(* IEC 61131-3 sources: sps-foerderband-sortieranlage/plc, 10 files *)

(* ---- E_Schritt.st ---- *)
{attribute 'qualified_only'}
{attribute 'strict'}
TYPE E_Schritt :
(
    INIT            := 0,   // Grundstellung herstellen
    BEREIT          := 1,   // Stillstand, wartet auf Start
    WARTEN_AUF_TEIL := 2,   // Automatik, wartet auf Teil an B1
    TRANSPORT       := 3,   // Band läuft, Material wird an B2 erkannt
    AUSWERFER_AUS   := 4,   // Metallteil: Auswerfer fährt aus
    AUSWERFER_EIN   := 5,   // Auswerfer fährt zurück
    STOERUNG        := 9    // Not-Halt oder Zeitüberschreitung
);
END_TYPE

(* ---- GVL_IO.st ---- *)
{attribute 'qualified_only'}
VAR_GLOBAL
    // ---------- Eingänge ----------
    // Öffner: TRUE = in Ordnung. Startwert TRUE nur für die Simulation,
    // weil es keinen realen Taster gibt, der den Kontakt geschlossen hält.
    xNotHaltOk            : BOOL := TRUE;   // S0  %IX0.0  Öffner
    xStart                : BOOL;           // S1  %IX0.1  Schließer
    xStoppOk              : BOOL := TRUE;   // S2  %IX0.2  Öffner
    xQuittieren           : BOOL;           // S3  %IX0.3  Schließer
    xZaehlerReset         : BOOL;           // S4  %IX0.4  Schließer
    xTeilEinlauf          : BOOL;           // B1  %IX0.5
    xTeilMetall           : BOOL;           // B2  %IX0.6  induktiv
    xTeilAuswurfPos       : BOOL;           // B3  %IX0.7
    xTeilRutscheB         : BOOL;           // B4  %IX1.0
    xAuswerferEingefahren : BOOL := TRUE;   // B5  %IX1.1
    xAuswerferAusgefahren : BOOL;           // B6  %IX1.2

    // ---------- Ausgänge ----------
    xBandMotor            : BOOL;           // K1/M1 %QX0.0
    xAuswerferAusfahren   : BOOL;           // Y1    %QX0.1
    xLampeBetrieb         : BOOL;           // H1    %QX0.2
    xLampeStoerung        : BOOL;           // H2    %QX0.3
END_VAR

(* ---- GVL_Param.st ---- *)
{attribute 'qualified_only'}
VAR_GLOBAL CONSTANT
    tTimeoutTransport : TIME := T#8S;     // Teil muss B3 bzw. B4 innerhalb dieser Zeit erreichen
    tTimeoutAuswerfer : TIME := T#2S;     // Auswerfer muss seine Endlage innerhalb dieser Zeit erreichen
    tBlinkHalbperiode : TIME := T#500MS;  // Blinktakt der Störungsleuchte
END_VAR

(* ---- GVL_Sim.st ---- *)
{attribute 'qualified_only'}
VAR_GLOBAL
    // ---------- Bedienung der Simulation (Visualisierung) ----------
    xMetallteilAuflegen     : BOOL;
    xKunststoffteilAuflegen : BOOL;
    xBandLeeren             : BOOL;      // Bediener nimmt ein Teil vom Band (z. B. nach Not-Halt)
    xZylinderKlemmt         : BOOL;      // Fehlersimulation: Auswerfer bewegt sich nicht

    // ---------- Zustand der Simulation (nur Anzeige) ----------
    xTeilAufBand            : BOOL;
    rTeilPosition           : REAL;      // mm ab Bandanfang
    rAuswerferPosition      : REAL;      // 0 = eingefahren, 100 = ausgefahren
END_VAR

(* ---- GVL_Status.st ---- *)
{attribute 'qualified_only'}
VAR_GLOBAL
    // ---------- Zustand (wird per OPC UA bereitgestellt) ----------
    eSchritt            : E_Schritt := E_Schritt.INIT;
    sSchritt            : STRING(30);
    xBetrieb            : BOOL;          // Automatikablauf aktiv
    xStoerung           : BOOL;          // Störung gespeichert, noch nicht quittiert
    xNotHaltAktiv       : BOOL;          // Not-Halt steht aktuell an
    sStoerung           : STRING(80);    // Störungstext

    // ---------- Zähler und Kennzahlen ----------
    uiAnzahlMetall      : UINT;
    uiAnzahlKunststoff  : UINT;
    uiAnzahlGesamt      : UINT;
    uiAnzahlNotHalt     : UINT;
    tLetzteZykluszeit   : TIME;          // Zeit vom Einlauf bis zum Abschluss des letzten Teils
    tStillstandGesamt   : TIME;          // aufsummierte Zeit im Störungszustand

    // ---------- interne Anforderungen Ablauf -> Ausgaben ----------
    xBandEin            : BOOL;
    xAuswerferEin       : BOOL;
END_VAR

(* ---- FB_Anlagensimulation.st ---- *)
FUNCTION_BLOCK FB_Anlagensimulation
VAR
    fbMetallFlanke     : R_TRIG;
    fbKunststoffFlanke : R_TRIG;
    fbLeerenFlanke     : R_TRIG;
    fbRutscheBImpuls   : TP;
    xTeilIstMetall     : BOOL;
    xTeilFaelltInB     : BOOL;
    xErsterZyklus      : BOOL := TRUE;
    tJetzt             : TIME;
    tLetzter           : TIME;
    rDt                : REAL;          // Zeit seit dem letzten Zyklus in s
END_VAR
VAR CONSTANT
    rBandGeschw        : REAL := 200.0;  // mm/s
    rBandLaenge        : REAL := 1000.0; // mm
    rB1Start           : REAL := 0.0;
    rB1Ende            : REAL := 80.0;
    rB2Start           : REAL := 350.0;
    rB2Ende            : REAL := 420.0;
    rB3Start           : REAL := 650.0;
    rB3Ende            : REAL := 720.0;
    rAuswerferGeschw   : REAL := 200.0;  // %/s, ein Hub dauert 0,5 s
    rAuswurfSchwelle   : REAL := 50.0;   // ab hier ist das Teil vom Band geschoben
END_VAR

(* ---------- Implementierung ---------- *)

// Zeitschritt bestimmen (begrenzt, damit Pausen im Debugger keine Sprünge erzeugen)
tJetzt := TIME();
IF xErsterZyklus THEN
    tLetzter := tJetzt;
    xErsterZyklus := FALSE;
END_IF
rDt := MIN(TIME_TO_REAL(tJetzt - tLetzter) / 1000.0, 0.1);
tLetzter := tJetzt;

// Teile auflegen und entfernen
fbMetallFlanke(CLK := GVL_Sim.xMetallteilAuflegen);
fbKunststoffFlanke(CLK := GVL_Sim.xKunststoffteilAuflegen);
fbLeerenFlanke(CLK := GVL_Sim.xBandLeeren);

IF NOT GVL_Sim.xTeilAufBand THEN
    IF fbMetallFlanke.Q THEN
        GVL_Sim.xTeilAufBand := TRUE;
        GVL_Sim.rTeilPosition := 0.0;
        xTeilIstMetall := TRUE;
    ELSIF fbKunststoffFlanke.Q THEN
        GVL_Sim.xTeilAufBand := TRUE;
        GVL_Sim.rTeilPosition := 0.0;
        xTeilIstMetall := FALSE;
    END_IF
END_IF

IF fbLeerenFlanke.Q THEN
    GVL_Sim.xTeilAufBand := FALSE;
END_IF

// Bandbewegung
xTeilFaelltInB := FALSE;
IF GVL_Sim.xTeilAufBand AND GVL_IO.xBandMotor THEN
    GVL_Sim.rTeilPosition := GVL_Sim.rTeilPosition + rBandGeschw * rDt;
    IF GVL_Sim.rTeilPosition >= rBandLaenge THEN
        GVL_Sim.xTeilAufBand := FALSE;
        xTeilFaelltInB := TRUE;
    END_IF
END_IF
fbRutscheBImpuls(IN := xTeilFaelltInB, PT := T#500MS);

// Auswerfer (bei Fehlersimulation bleibt er stehen)
IF NOT GVL_Sim.xZylinderKlemmt THEN
    IF GVL_IO.xAuswerferAusfahren THEN
        GVL_Sim.rAuswerferPosition := MIN(GVL_Sim.rAuswerferPosition + rAuswerferGeschw * rDt, 100.0);
    ELSE
        GVL_Sim.rAuswerferPosition := MAX(GVL_Sim.rAuswerferPosition - rAuswerferGeschw * rDt, 0.0);
    END_IF
END_IF

// Auswurf in Rutsche A
IF GVL_Sim.xTeilAufBand
   AND GVL_Sim.rAuswerferPosition >= rAuswurfSchwelle
   AND GVL_Sim.rTeilPosition >= rB3Start
   AND GVL_Sim.rTeilPosition <= rB3Ende THEN
    GVL_Sim.xTeilAufBand := FALSE;
END_IF

// Sensorsignale
GVL_IO.xTeilEinlauf := GVL_Sim.xTeilAufBand
                       AND GVL_Sim.rTeilPosition >= rB1Start
                       AND GVL_Sim.rTeilPosition <= rB1Ende;
GVL_IO.xTeilMetall := GVL_Sim.xTeilAufBand AND xTeilIstMetall
                      AND GVL_Sim.rTeilPosition >= rB2Start
                      AND GVL_Sim.rTeilPosition <= rB2Ende;
GVL_IO.xTeilAuswurfPos := GVL_Sim.xTeilAufBand
                          AND GVL_Sim.rTeilPosition >= rB3Start
                          AND GVL_Sim.rTeilPosition <= rB3Ende;
GVL_IO.xTeilRutscheB := fbRutscheBImpuls.Q;
GVL_IO.xAuswerferEingefahren := GVL_Sim.rAuswerferPosition <= 0.5;
GVL_IO.xAuswerferAusgefahren := GVL_Sim.rAuswerferPosition >= 99.5;

(* ---- PLC_PRG.st ---- *)
PROGRAM PLC_PRG
VAR
    fbAnlage : FB_Anlagensimulation;
END_VAR

(* ---------- Implementierung ---------- *)

// Reihenfolge: Sensoren erzeugen, Störungen auswerten, Ablauf, Ausgänge schreiben
fbAnlage();
PRG_Stoerung();
PRG_Ablauf();
PRG_Ausgaben();

(* ---- PRG_Ablauf.st ---- *)
PROGRAM PRG_Ablauf
VAR
    fbStartFlanke     : R_TRIG;
    fbResetFlanke     : R_TRIG;
    fbSchrittZeit     : TON;                       // misst, wie lange der aktuelle Schritt schon aktiv ist
    eSchrittAlt       : E_Schritt := E_Schritt.INIT;
    xStoppAngefordert : BOOL;                      // Stopp am Zyklusende
    xIstMetall        : BOOL;                      // an B2 erkanntes Material des aktuellen Teils
    tTeilStart        : TIME;
END_VAR

(* ---------- Implementierung ---------- *)

fbStartFlanke(CLK := GVL_IO.xStart);
fbResetFlanke(CLK := GVL_IO.xZaehlerReset);

// Schrittzeit: wird bei jedem Schrittwechsel für einen Zyklus zurückgesetzt
fbSchrittZeit(IN := (GVL_Status.eSchritt = eSchrittAlt), PT := T#24H);
eSchrittAlt := GVL_Status.eSchritt;

// Stopp (Öffner) nur merken, das aktuelle Teil wird fertig bearbeitet
IF NOT GVL_IO.xStoppOk THEN
    xStoppAngefordert := TRUE;
END_IF

// Eine Störung hat Vorrang vor jedem Schritt
IF GVL_Status.xStoerung THEN
    GVL_Status.eSchritt := E_Schritt.STOERUNG;
END_IF

CASE GVL_Status.eSchritt OF

    E_Schritt.INIT:
        GVL_Status.xBandEin := FALSE;
        GVL_Status.xAuswerferEin := FALSE;
        IF GVL_IO.xAuswerferEingefahren THEN
            GVL_Status.eSchritt := E_Schritt.BEREIT;
        ELSIF fbSchrittZeit.ET > GVL_Param.tTimeoutAuswerfer THEN
            GVL_Status.xStoerung := TRUE;
            GVL_Status.sStoerung := 'Grundstellung: Auswerfer faehrt nicht ein (B5)';
            GVL_Status.eSchritt := E_Schritt.STOERUNG;
        END_IF

    E_Schritt.BEREIT:
        GVL_Status.xBandEin := FALSE;
        GVL_Status.xAuswerferEin := FALSE;
        IF fbResetFlanke.Q THEN
            GVL_Status.uiAnzahlMetall := 0;
            GVL_Status.uiAnzahlKunststoff := 0;
            GVL_Status.uiAnzahlGesamt := 0;
        END_IF
        // Wiederanlaufsperre: Start nur mit neuer Flanke
        IF fbStartFlanke.Q AND GVL_IO.xStoppOk THEN
            xStoppAngefordert := FALSE;
            GVL_Status.eSchritt := E_Schritt.WARTEN_AUF_TEIL;
        END_IF

    E_Schritt.WARTEN_AUF_TEIL:
        GVL_Status.xBandEin := FALSE;
        GVL_Status.xAuswerferEin := FALSE;
        IF xStoppAngefordert THEN
            GVL_Status.eSchritt := E_Schritt.BEREIT;
        ELSIF GVL_IO.xTeilEinlauf THEN
            xIstMetall := FALSE;
            tTeilStart := TIME();
            GVL_Status.eSchritt := E_Schritt.TRANSPORT;
        END_IF

    E_Schritt.TRANSPORT:
        GVL_Status.xBandEin := TRUE;
        GVL_Status.xAuswerferEin := FALSE;
        // Das Signal von B2 ist nur kurz da, deshalb wird das Material gespeichert
        IF GVL_IO.xTeilMetall THEN
            xIstMetall := TRUE;
        END_IF
        IF xIstMetall AND GVL_IO.xTeilAuswurfPos THEN
            GVL_Status.xBandEin := FALSE;
            GVL_Status.eSchritt := E_Schritt.AUSWERFER_AUS;
        ELSIF NOT xIstMetall AND GVL_IO.xTeilRutscheB THEN
            GVL_Status.xBandEin := FALSE;
            GVL_Status.uiAnzahlKunststoff := GVL_Status.uiAnzahlKunststoff + 1;
            GVL_Status.uiAnzahlGesamt := GVL_Status.uiAnzahlGesamt + 1;
            GVL_Status.tLetzteZykluszeit := TIME() - tTeilStart;
            IF xStoppAngefordert THEN
                GVL_Status.eSchritt := E_Schritt.BEREIT;
            ELSE
                GVL_Status.eSchritt := E_Schritt.WARTEN_AUF_TEIL;
            END_IF
        ELSIF fbSchrittZeit.ET > GVL_Param.tTimeoutTransport THEN
            GVL_Status.xStoerung := TRUE;
            GVL_Status.sStoerung := 'Transport: Teil erreicht B3 bzw. B4 nicht';
            GVL_Status.eSchritt := E_Schritt.STOERUNG;
        END_IF

    E_Schritt.AUSWERFER_AUS:
        GVL_Status.xBandEin := FALSE;
        GVL_Status.xAuswerferEin := TRUE;
        IF GVL_IO.xAuswerferAusgefahren THEN
            GVL_Status.eSchritt := E_Schritt.AUSWERFER_EIN;
        ELSIF fbSchrittZeit.ET > GVL_Param.tTimeoutAuswerfer THEN
            GVL_Status.xStoerung := TRUE;
            GVL_Status.sStoerung := 'Auswerfer erreicht vordere Endlage nicht (B6)';
            GVL_Status.eSchritt := E_Schritt.STOERUNG;
        END_IF

    E_Schritt.AUSWERFER_EIN:
        GVL_Status.xBandEin := FALSE;
        GVL_Status.xAuswerferEin := FALSE;
        IF GVL_IO.xAuswerferEingefahren THEN
            GVL_Status.uiAnzahlMetall := GVL_Status.uiAnzahlMetall + 1;
            GVL_Status.uiAnzahlGesamt := GVL_Status.uiAnzahlGesamt + 1;
            GVL_Status.tLetzteZykluszeit := TIME() - tTeilStart;
            IF xStoppAngefordert THEN
                GVL_Status.eSchritt := E_Schritt.BEREIT;
            ELSE
                GVL_Status.eSchritt := E_Schritt.WARTEN_AUF_TEIL;
            END_IF
        ELSIF fbSchrittZeit.ET > GVL_Param.tTimeoutAuswerfer THEN
            GVL_Status.xStoerung := TRUE;
            GVL_Status.sStoerung := 'Auswerfer erreicht hintere Endlage nicht (B5)';
            GVL_Status.eSchritt := E_Schritt.STOERUNG;
        END_IF

    E_Schritt.STOERUNG:
        GVL_Status.xBandEin := FALSE;
        GVL_Status.xAuswerferEin := FALSE;
        // Nach dem Quittieren zurück in die Grundstellung, danach ist ein neuer Start nötig
        IF NOT GVL_Status.xStoerung THEN
            GVL_Status.eSchritt := E_Schritt.INIT;
        END_IF

END_CASE

// Anzeige und Betriebsstatus
GVL_Status.xBetrieb := GVL_Status.eSchritt = E_Schritt.WARTEN_AUF_TEIL
                       OR GVL_Status.eSchritt = E_Schritt.TRANSPORT
                       OR GVL_Status.eSchritt = E_Schritt.AUSWERFER_AUS
                       OR GVL_Status.eSchritt = E_Schritt.AUSWERFER_EIN;

CASE GVL_Status.eSchritt OF
    E_Schritt.INIT:            GVL_Status.sSchritt := 'Grundstellung';
    E_Schritt.BEREIT:          GVL_Status.sSchritt := 'Bereit';
    E_Schritt.WARTEN_AUF_TEIL: GVL_Status.sSchritt := 'Warten auf Teil';
    E_Schritt.TRANSPORT:       GVL_Status.sSchritt := 'Transport';
    E_Schritt.AUSWERFER_AUS:   GVL_Status.sSchritt := 'Auswerfer faehrt aus';
    E_Schritt.AUSWERFER_EIN:   GVL_Status.sSchritt := 'Auswerfer faehrt ein';
    E_Schritt.STOERUNG:        GVL_Status.sSchritt := 'Stoerung';
END_CASE

(* ---- PRG_Ausgaben.st ---- *)
PROGRAM PRG_Ausgaben
VAR
    fbBlinkTakt : TON;
    xBlink      : BOOL;
    xFreigabe   : BOOL;
END_VAR

(* ---------- Implementierung ---------- *)

// Aktoren nur bei entriegeltem Not-Halt und ohne Störung freigeben
xFreigabe := GVL_IO.xNotHaltOk AND NOT GVL_Status.xStoerung;

GVL_IO.xBandMotor          := GVL_Status.xBandEin AND xFreigabe;
GVL_IO.xAuswerferAusfahren := GVL_Status.xAuswerferEin AND xFreigabe;   // FALSE: Federrückstellung fährt ein
GVL_IO.xLampeBetrieb       := GVL_Status.xBetrieb AND xFreigabe;

// Störungsleuchte: Dauerlicht solange der Not-Halt ansteht, Blinken bis zur Quittierung
fbBlinkTakt(IN := NOT fbBlinkTakt.Q, PT := GVL_Param.tBlinkHalbperiode);
IF fbBlinkTakt.Q THEN
    xBlink := NOT xBlink;
END_IF

IF GVL_Status.xNotHaltAktiv THEN
    GVL_IO.xLampeStoerung := TRUE;
ELSIF GVL_Status.xStoerung THEN
    GVL_IO.xLampeStoerung := xBlink;
ELSE
    GVL_IO.xLampeStoerung := FALSE;
END_IF

(* ---- PRG_Stoerung.st ---- *)
PROGRAM PRG_Stoerung
VAR
    fbNotHaltFlanke : R_TRIG;   // Not-Halt wurde betätigt (für den Ereigniszähler)
    fbQuittFlanke   : R_TRIG;
    tJetzt          : TIME;
    tLetzter        : TIME;
END_VAR

(* ---------- Implementierung ---------- *)

tJetzt := TIME();

// Not-Halt (Öffner): FALSE bedeutet betätigt oder Leitungsbruch
GVL_Status.xNotHaltAktiv := NOT GVL_IO.xNotHaltOk;

fbNotHaltFlanke(CLK := GVL_Status.xNotHaltAktiv);
IF fbNotHaltFlanke.Q THEN
    GVL_Status.uiAnzahlNotHalt := GVL_Status.uiAnzahlNotHalt + 1;
END_IF

// Solange der Not-Halt ansteht, bleibt die Störung gesetzt
IF GVL_Status.xNotHaltAktiv THEN
    GVL_Status.xStoerung := TRUE;
    GVL_Status.sStoerung := 'Not-Halt betaetigt';
END_IF

// Quittieren nur mit neuer Flanke und nur, wenn der Not-Halt entriegelt ist.
// Zeitüberschreitungen setzt PRG_Ablauf direkt in GVL_Status.
fbQuittFlanke(CLK := GVL_IO.xQuittieren);
IF fbQuittFlanke.Q AND GVL_Status.xStoerung AND GVL_IO.xNotHaltOk THEN
    GVL_Status.xStoerung := FALSE;
    GVL_Status.sStoerung := '';
END_IF

// Stillstandszeit für die Kennzahlen aufsummieren
IF GVL_Status.xStoerung THEN
    GVL_Status.tStillstandGesamt := GVL_Status.tStillstandGesamt + (tJetzt - tLetzter);
END_IF
tLetzter := tJetzt;
